(* IEC 61131-3 sources: st2fb/corpus/00_latch, 1 file *)

(* ---- program.st ---- *)
FUNCTION_BLOCK LATCH
VAR_INPUT
  S : BOOL;
  R : BOOL;
END_VAR
VAR_OUTPUT
  Q : BOOL;
  COUNT : INT;
END_VAR
VAR
  PREV : BOOL;
END_VAR
  IF R THEN
    Q := FALSE;
  ELSIF S THEN
    Q := TRUE;
  END_IF;
  IF Q AND NOT PREV THEN
    COUNT := COUNT + 1;
  END_IF;
  PREV := Q;
END_FUNCTION_BLOCK
